(* IEC 61131-3 sources: rusty/tests/lit/cfc/generics/generic_chain, 2 files *)

(* ---- main.st ---- *)
FUNCTION main : DINT
    generic_chain.a := 1000;
    generic_chain.b := 2000;
    generic_chain.c := 100000;
    generic_chain();
    // CHECK: result = 103000
    printf('result = %d$N', generic_chain.result);
END_FUNCTION

(* ---- myGenAdd.st ---- *)
FUNCTION myGenAdd<T: ANY_NUM> : T
VAR_INPUT
    a : T;
    b : T;
END_VAR
END_FUNCTION

FUNCTION myGenAdd__INT : INT
VAR_INPUT
    a : INT;
    b : INT;
END_VAR
    myGenAdd__INT := a + b;
END_FUNCTION

FUNCTION myGenAdd__DINT : DINT
VAR_INPUT
    a : DINT;
    b : DINT;
END_VAR
    myGenAdd__DINT := a + b;
END_FUNCTION
